(* IEC 61131-3 sources: llm-plc-st-eval/data/processed_definitivo/gemini-3.1-pro-preview/C3/few_shot, 3 files *)

(* ---- ejec_1.st ---- *)
PROGRAM PRG_Conversion
VAR_INPUT
    btnMarcha : BOOL; (* Contacto NA en paralelo con motor *)
    btnParo : BOOL; (* Contacto NC en serie *)
END_VAR
VAR_OUTPUT
    motor : BOOL; (* Bobina y contacto de retencion *)
    lampara : BOOL; (* Bobina activada por el temporizador *)
END_VAR
VAR
    T1 : TON; (* Temporizador a la conexion *)
END_VAR

(* Rama 1: Circuito de marcha/paro con auto-retencion *)
motor := (btnMarcha OR motor) AND NOT btnParo;

(* Rama 2: Temporizador alimentado por el estado del motor *)
T1(IN := motor, PT := T#10S);

(* Rama 3: Activacion de la lampara con la salida del temporizador *)
lampara := T1.Q;
END_PROGRAM

(* ---- ejec_2.st ---- *)
PROGRAM PRG_Conversion
VAR_INPUT
    btnMarcha : BOOL; (* Contacto NA, inicio de marcha *)
    btnParo : BOOL; (* Contacto NC, detiene el motor *)
END_VAR
VAR_OUTPUT
    motor : BOOL; (* Bobina del motor y contacto de retencion *)
    lampara : BOOL; (* Bobina indicadora *)
END_VAR
VAR
    T1 : TON; (* Temporizador a la conexion *)
END_VAR

(* Rama 1: Circuito de retencion (arranque/paro) para el motor *)
motor := (btnMarcha OR motor) AND NOT btnParo;

(* Rama 2: El temporizador se activa cuando el motor esta encendido *)
T1(IN := motor, PT := T#10S);

(* Rama 3: La lampara se enciende cuando el temporizador alcanza los 10s *)
lampara := T1.Q;
END_PROGRAM

(* ---- ejec_3.st ---- *)
PROGRAM PRG_Conversion
VAR_INPUT
    btnMarcha : BOOL; (* Contacto NA en paralelo *)
    btnParo : BOOL; (* Contacto NC en serie *)
END_VAR
VAR_OUTPUT
    motor : BOOL; (* Bobina y contacto NA de realimentacion *)
    lampara : BOOL; (* Bobina indicadora *)
END_VAR
VAR
    T1 : TON; (* Temporizador a la conexion *)
END_VAR

(* Rama 1: Arranque y paro del motor con auto-retencion *)
motor := (btnMarcha OR motor) AND NOT btnParo;

(* Rama 2: Temporizador de 10 segundos activado por el motor *)
T1(IN := motor, PT := T#10S);

(* Rama 3: Activacion de la lampara con la salida del temporizador *)
lampara := T1.Q;
END_PROGRAM
